(* Schneider Machine Expert - Basic project timer_profile_02_10ms_all, file version 3.0.0.0 *)
(* ProjectInformations: Name=New project *)

HARDWARE
  Cpu 0: TM200CE40T
  EthernetConfiguration: NetworkName=M200, IpAllocationMode=FixedAddress, IpAddress=0.0.0.0, SubnetMask=0.0.0.0
  SerialLineConfiguration: Baud=Baud19200, Parity=ParityEven, DataBits=DataBits8, StopBits=StopBits1, PhysicalMedium=PhysicalMediumRs485, TransmissionMode=TransmissionModeModbusRtu, SlaveId=1, Addressing=SlaveAddressing
  MastTask: UsePeriodScanMode=false, PeriodScan=100
  FastTask: Period=255
  CpuBehavior: StartingMode=StartAsPreviousState, AutoSaveRamOnEeprom=true, WatchdogPeriod=250

SYMBOLS  (address, symbol, comment, settings)
  %TM0        [Preset=5, Base=TenMilliSeconds]
  %TM1        [Type=TOF, Preset=5, Base=TenMilliSeconds]
  %TM2        [Type=TP, Preset=5, Base=TenMilliSeconds]

POU New POU
  (* SectionNumber=0 *)

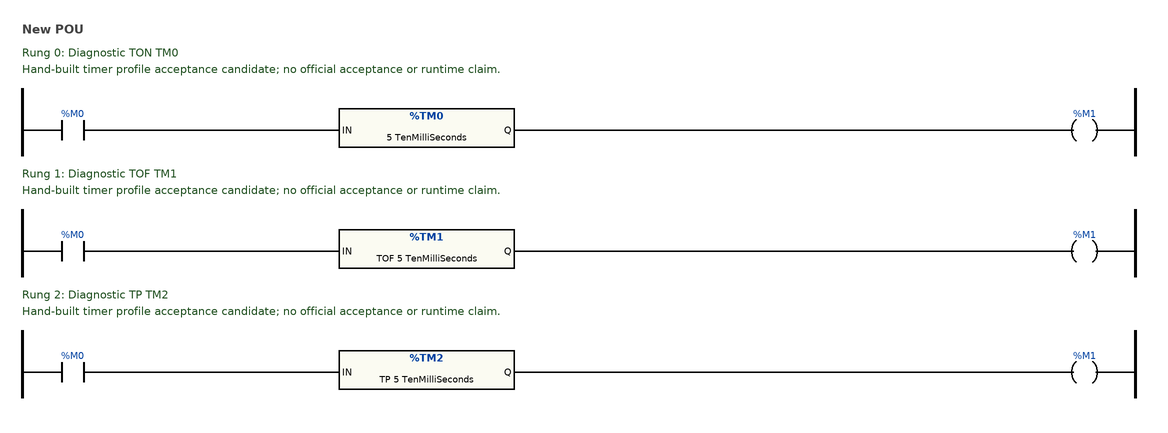

// Rung 0: Diagnostic TON TM0
// Hand-built timer profile acceptance candidate; no official acceptance or runtime claim.
  BLK %TM0
  LD %M0
  IN
  OUT_BLK
  LD Q
  ST %M1
  END_BLK
  // as ST:
  //   %TM0(IN := %M0);
  //   %M1 := %TM0.Q;

// Rung 1: Diagnostic TOF TM1
// Hand-built timer profile acceptance candidate; no official acceptance or runtime claim.
  BLK %TM1
  LD %M0
  IN
  OUT_BLK
  LD Q
  ST %M1
  END_BLK
  // as ST:
  //   %TM1(IN := %M0);
  //   %M1 := %TM1.Q;

// Rung 2: Diagnostic TP TM2
// Hand-built timer profile acceptance candidate; no official acceptance or runtime claim.
  BLK %TM2
  LD %M0
  IN
  OUT_BLK
  LD Q
  ST %M1
  END_BLK
  // as ST:
  //   %TM2(IN := %M0);
  //   %M1 := %TM2.Q;
